Fanuc KAREL source: KB00071.KL

PROGRAM KB00071
%NOLOCKGROUP
VAR
  P1: REAL
  RESULT: REAL
BEGIN
  P1 = 1.0
  RESULT = EXP(P1)
END KB00071
